Universal Robots URScript: T006_codellama_34b_adversarial_A8.5_rep1.urscript

def bin_picking():
    # Home position
    movej(p[0, 0, 0, 0, 0, 0], v=350.0)

    # Above bin
    movel(p[0, 0, 120, 0, 0, 0], v=350.0)

    # Descend
